// TIA Portal V21 export
// export: Created 2026-11-07T14:35:59.5082391Z, ExportSetting WithDefaults, DisplayName Totally Integrated Automation Portal, DisplayVersion V21, DisplayName STEP 7 Professional, DisplayVersion V21, DisplayName STEP 7 Safety, DisplayVersion V21, DisplayName Tech WebApplication, DisplayVersion V21, DisplayName WinCC Basic/Comfort/Advanced, DisplayVersion V21, DisplayName WinCC Unified, DisplayVersion V21
Screen "T12_DT"  1024x768, Number=32
  ScreenLayer 
    DateTimeField "P_DateTime" at 10,10 size 346x40  Mode=Output
